{attribute 'no_assign'}
FUNCTION_BLOCK FB_DO_WTURBINE_LD0_WPPD1_ClrOp EXTENDS FB_AcsiCommonDataClass
VAR_INPUT
	st_: FB_DO_WTURBINE_LD0_WPPD1_ClrOp_st := (sObjectName:='st', sClass:='ENC', bLinkResult:=THIS^.AddDataToContainer(ipData:=st_));
END_VAR
VAR
END_VAR

END_FUNCTION_BLOCK

(* stored: Version 1.1.0.1
   POU FB_DO_WTURBINE_LD0_WPPD1_ClrOp: Id {6d9b2bcf-91b9-448d-9934-175eeced678f}, SpecialFunc None *)
